// TIA Portal V17 export
// export: Created 2026-11-10T15:00:48.6641979Z, ExportSetting WithDefaults, DisplayName Totally Integrated Automation Portal, DisplayVersion V17, DisplayName TIA Portal Openness, DisplayVersion V17, DisplayName TIA Portal Version Control Interface, DisplayVersion V17, DisplayName STEP 7 Professional, DisplayVersion V17, DisplayName STEP 7 Safety, DisplayVersion V17, DisplayName WinCC Advanced, DisplayVersion V17
GraphicList "Level150"  ListRange=Decimal, Mode=Simple
  GraphicListEntry   EntryType=Range, To=14, Picture=Tank_0
  GraphicListEntry   EntryType=Range, From=15, To=29, Picture=Tank_1
  GraphicListEntry   EntryType=Range, From=30, To=44, Picture=Tank_2
  GraphicListEntry   EntryType=Range, From=45, To=59, Picture=Tank_3
  GraphicListEntry   EntryType=Range, From=60, To=74, Picture=Tank_4
  GraphicListEntry   EntryType=Range, From=75, To=89, Picture=Tank_5
  GraphicListEntry   EntryType=Range, From=90, To=104, Picture=Tank_6
  GraphicListEntry   EntryType=Range, From=105, To=119, Picture=Tank_7
  GraphicListEntry   EntryType=Range, From=120, To=134, Picture=Tank_8
  GraphicListEntry   EntryType=Range, From=135, To=149, Picture=Tank_9
  GraphicListEntry   EntryType=Range, From=150, To=150, Picture=Tank_10
